Universal Robots URScript: SF1_Rotation_17_Sequence.script

# Case 17 of sf1_plc_v4.script, the rotation sequence home -> home, optimised: the station lines
# verbatim from the program, the transfer segments S1-S3 generated movej (the program's a and v,
# r=0). Points: SF1_Rotation_17.urscript.
# The station lines to Waypoint_4, Waypoint_5, pick_rotate_1, Waypoint_6 are the program's text; their points have the program's _p and
# another _q (SF1_Rotation_17.urscript).
# Machine margin: generated segments keep 30.0 mm (Clearance.Environment 20.0 + Machine_Extra 10.0 mm) to machine_a
# outside the station zone; source: owner accuracy estimate of the machine position, 2026-10-18.
# Variant c2: delivered - tested on the real cell (owner, 2026-10-21), = Data/Generated/: the drop on branch S- E- W- (wrist flipped in S1).
# Simulation passed != safe on the robot: run it at reduced speed first.
# Start at home (generated, r=0): the program's line blends (r=0.01) into S1, and a blend into a generated segment is not checked
movej(home_q, a=1.3962634015954636, v=1.0471975511965976, r=0)
# S1 (generated): home -> drop_rotate_1
movej(drop_rotate_1_q, a=1.3962634015954636, v=1.0471975511965976, r=0)
# Station: drop (verbatim from the program)
movel(Waypoint_4_p, a=1.2, v=0.25)
# Gripper open: the program's Robotiq node goes here (rq_set_pos_spd_for(0, 255, 255, "1"))
movej(get_inverse_kin(Waypoint_5_p, qnear=Waypoint_5_q), a=1.3962634015954636, v=1.0471975511965976)
# S2 (generated): Waypoint_5 -> Waypoint_18
movej(via_Waypoint_5_Waypoint_18_01_q, a=1.3962634015954636, v=1.0471975511965976, r=0)
movej(Waypoint_18_q, a=1.3962634015954636, v=1.0471975511965976, r=0)
# Station: pick (verbatim from the program)
movej(get_inverse_kin(pick_rotate_1_p, qnear=pick_rotate_1_q), a=1.3962634015954636, v=1.0471975511965976)
# Gripper close: the program's Robotiq node goes here (rq_set_pos_spd_for(255, 255, 255, "1"))
movel(Waypoint_6_p, a=1.2, v=0.25)
# S3 (generated): Waypoint_6 -> home
movej(via_Waypoint_6_home_01_q, a=1.3962634015954636, v=1.0471975511965976, r=0)
movej(home_q, a=1.3962634015954636, v=1.0471975511965976, r=0)
